FUNCTION_BLOCK UV_Trojan_HMI (* Service Interface Function Block Type *)
  (* Standard: 61499-2 *)
  (* Version 1.0, 19/10/2026, Hidryco, Hidryco, IHM do UV_Trojan *)
  PACKAGE Hidryco.HidrycoLib;
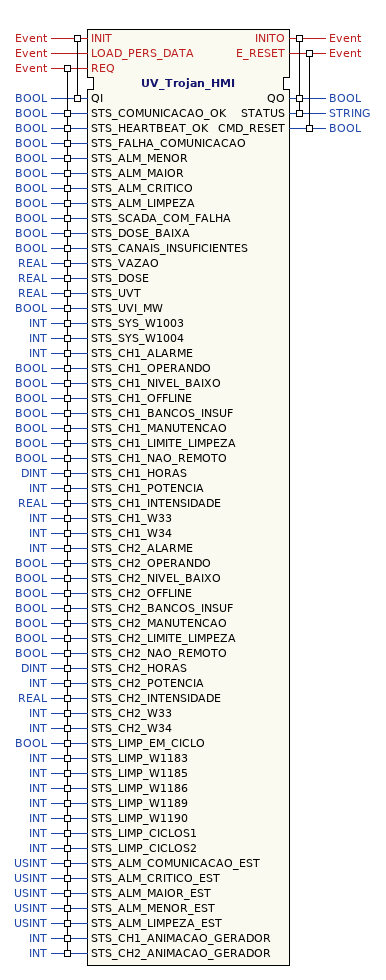
  EVENT_INPUT
    INIT WITH QI;
    LOAD_PERS_DATA; (* Reenvia os parametros persistentes *)
    REQ WITH STS_COMUNICACAO_OK, STS_HEARTBEAT_OK, STS_FALHA_COMUNICACAO, STS_ALM_MENOR, STS_ALM_MAIOR, STS_ALM_CRITICO, STS_ALM_LIMPEZA, STS_SCADA_COM_FALHA, STS_DOSE_BAIXA, STS_CANAIS_INSUFICIENTES, STS_VAZAO, STS_DOSE, STS_UVT, STS_UVI_MW, STS_SYS_W1003, STS_SYS_W1004, STS_CH1_ALARME, STS_CH1_OPERANDO, STS_CH1_NIVEL_BAIXO, STS_CH1_OFFLINE, STS_CH1_BANCOS_INSUF, STS_CH1_MANUTENCAO, STS_CH1_LIMITE_LIMPEZA, STS_CH1_NAO_REMOTO, STS_CH1_HORAS, STS_CH1_POTENCIA, STS_CH1_INTENSIDADE, STS_CH1_W33, STS_CH1_W34, STS_CH2_ALARME, STS_CH2_OPERANDO, STS_CH2_NIVEL_BAIXO, STS_CH2_OFFLINE, STS_CH2_BANCOS_INSUF, STS_CH2_MANUTENCAO, STS_CH2_LIMITE_LIMPEZA, STS_CH2_NAO_REMOTO, STS_CH2_HORAS, STS_CH2_POTENCIA, STS_CH2_INTENSIDADE, STS_CH2_W33, STS_CH2_W34, STS_LIMP_EM_CICLO, STS_LIMP_W1183, STS_LIMP_W1185, STS_LIMP_W1186, STS_LIMP_W1189, STS_LIMP_W1190, STS_LIMP_CICLOS1, STS_LIMP_CICLOS2, STS_ALM_COMUNICACAO_EST, STS_ALM_CRITICO_EST, STS_ALM_MAIOR_EST, STS_ALM_MENOR_EST, STS_ALM_LIMPEZA_EST, STS_CH1_ANIMACAO_GERADOR, STS_CH2_ANIMACAO_GERADOR; (* Atualizacao de status *)
  END_EVENT
  EVENT_OUTPUT
    INITO WITH QO, STATUS;
    E_RESET WITH CMD_RESET;
  END_EVENT
  VAR_INPUT
    QI : BOOL;
    STS_COMUNICACAO_OK : BOOL; (* Comunicacao Modbus e heartbeat do SCC OK *)
    STS_HEARTBEAT_OK : BOOL; (* Heartbeat do SCC (41001.8) alternando *)
    STS_FALHA_COMUNICACAO : BOOL; (* Falha de comunicacao com o SCC *)
    STS_ALM_MENOR : BOOL; (* Alarme comum menor (41001.0) *)
    STS_ALM_MAIOR : BOOL; (* Alarme comum maior (41001.1) *)
    STS_ALM_CRITICO : BOOL; (* Alarme comum critico (41001.2) *)
    STS_ALM_LIMPEZA : BOOL; (* Alarme do sistema de limpeza (41001.3) *)
    STS_SCADA_COM_FALHA : BOOL; (* SCC sem o heartbeat do CLP (41004.4) *)
    STS_DOSE_BAIXA : BOOL; (* Dose abaixo do alvo (41003.0) *)
    STS_CANAIS_INSUFICIENTES : BOOL; (* Canais saudaveis insuficientes (41003.1) *)
    STS_VAZAO : REAL; (* Vazao do sistema no SCC (41005 x fator 41008) *)
    STS_DOSE : REAL; (* Dose equivalente RED (mJ/cm2) *)
    STS_UVT : REAL; (* Transmitancia UV (%) *)
    STS_UVI_MW : BOOL; (* Unidade da intensidade: FALSE = %, TRUE = mW/cm2 *)
    STS_SYS_W1003 : INT; (* Registro 41003 (diagnostico) *)
    STS_SYS_W1004 : INT; (* Registro 41004 (diagnostico) *)
    STS_CH1_ALARME : INT; (* Canal 1: 0 normal, 1 menor, 2 maior, 3 critico *)
    STS_CH1_OPERANDO : BOOL; (* Canal 1 em operacao *)
    STS_CH1_NIVEL_BAIXO : BOOL; (* Canal 1 nivel de agua baixo *)
    STS_CH1_OFFLINE : BOOL; (* Canal 1 em modo offline *)
    STS_CH1_BANCOS_INSUF : BOOL; (* Canal 1 bancos saudaveis insuficientes *)
    STS_CH1_MANUTENCAO : BOOL; (* Canal 1 em manutencao *)
    STS_CH1_LIMITE_LIMPEZA : BOOL; (* Canal 1 vazao acima do limite de limpeza *)
    STS_CH1_NAO_REMOTO : BOOL; (* Banco do canal 1 fora de remoto automatico *)
    STS_CH1_HORAS : DINT; (* Banco do canal 1: horas das lampadas *)
    STS_CH1_POTENCIA : INT; (* Banco do canal 1: potencia (%) *)
    STS_CH1_INTENSIDADE : REAL; (* Banco do canal 1: intensidade UV *)
    STS_CH1_W33 : INT; (* Banco do canal 1: falhas 1 (diagnostico) *)
    STS_CH1_W34 : INT; (* Banco do canal 1: falhas 2 (diagnostico) *)
    STS_CH2_ALARME : INT; (* Canal 2: 0 normal, 1 menor, 2 maior, 3 critico *)
    STS_CH2_OPERANDO : BOOL; (* Canal 2 em operacao *)
    STS_CH2_NIVEL_BAIXO : BOOL; (* Canal 2 nivel de agua baixo *)
    STS_CH2_OFFLINE : BOOL; (* Canal 2 em modo offline *)
    STS_CH2_BANCOS_INSUF : BOOL; (* Canal 2 bancos saudaveis insuficientes *)
    STS_CH2_MANUTENCAO : BOOL; (* Canal 2 em manutencao *)
    STS_CH2_LIMITE_LIMPEZA : BOOL; (* Canal 2 vazao acima do limite de limpeza *)
    STS_CH2_NAO_REMOTO : BOOL; (* Banco do canal 2 fora de remoto automatico *)
    STS_CH2_HORAS : DINT; (* Banco do canal 2: horas das lampadas *)
    STS_CH2_POTENCIA : INT; (* Banco do canal 2: potencia (%) *)
    STS_CH2_INTENSIDADE : REAL; (* Banco do canal 2: intensidade UV *)
    STS_CH2_W33 : INT; (* Banco do canal 2: falhas 1 (diagnostico) *)
    STS_CH2_W34 : INT; (* Banco do canal 2: falhas 2 (diagnostico) *)
    STS_LIMP_EM_CICLO : BOOL; (* Sistema de limpeza em ciclo *)
    STS_LIMP_W1183 : INT; (* Registro 41183 (diagnostico) *)
    STS_LIMP_W1185 : INT; (* Registro 41185 (diagnostico) *)
    STS_LIMP_W1186 : INT; (* Registro 41186 (diagnostico) *)
    STS_LIMP_W1189 : INT; (* Registro 41189 (diagnostico) *)
    STS_LIMP_W1190 : INT; (* Registro 41190 (diagnostico) *)
    STS_LIMP_CICLOS1 : INT; (* Ciclos de limpeza do grupo 1 (canal 1) *)
    STS_LIMP_CICLOS2 : INT; (* Ciclos de limpeza do grupo 2 (canal 2) *)
    STS_ALM_COMUNICACAO_EST : USINT; (* Estado do ALARM_BIT (0 normal, 1 ativo reconhecido, 2 ativo nao reconhecido, 3 saiu nao reconhecido, 4 ativo e saiu nao reconhecido) *)
    STS_ALM_CRITICO_EST : USINT; (* Estado do ALARM_BIT (0 normal, 1 ativo reconhecido, 2 ativo nao reconhecido, 3 saiu nao reconhecido, 4 ativo e saiu nao reconhecido) *)
    STS_ALM_MAIOR_EST : USINT; (* Estado do ALARM_BIT (0 normal, 1 ativo reconhecido, 2 ativo nao reconhecido, 3 saiu nao reconhecido, 4 ativo e saiu nao reconhecido) *)
    STS_ALM_MENOR_EST : USINT; (* Estado do ALARM_BIT (0 normal, 1 ativo reconhecido, 2 ativo nao reconhecido, 3 saiu nao reconhecido, 4 ativo e saiu nao reconhecido) *)
    STS_ALM_LIMPEZA_EST : USINT; (* Estado do ALARM_BIT (0 normal, 1 ativo reconhecido, 2 ativo nao reconhecido, 3 saiu nao reconhecido, 4 ativo e saiu nao reconhecido) *)
    STS_CH1_ANIMACAO_GERADOR : INT; (* Raio do gerador do canal 1 (0..3) *)
    STS_CH2_ANIMACAO_GERADOR : INT; (* Raio do gerador do canal 2 (0..3) *)
  END_VAR
  VAR_OUTPUT
    QO : BOOL; (* Event Output Qualifier *)
    STATUS : STRING; (* Service Status *)
    CMD_RESET : BOOL; (* Reconhece os alarmes do UV *)
  END_VAR
  SERVICE /
    SEQUENCE 
    END_SEQUENCE
  END_SERVICE
END_FUNCTION_BLOCK
